(* IEC 61131-3 sources: 89152_FlorisHendrix_AfstudeerProject/89152_FlorisHendrix_ExamenProject/Stations/MachineControl/MachineControl/Class/VaranManager (part 5) *)

                DPRAM_Used.Total  += TempMem;
                DOCounter.Total   += 1;

            VARAN_CMD_CONTROL_WRITE,
            VARAN_CMD_MEMORY_WRITE:     // Write DO -------------------------------------------------------------------------------------------------------------------------------
                //32 Byte (Header) + 6 Byte (1 Byte Cmd, 4 Byte Addr, 1 Byte Len) + 1 Byte (Response) + n Byte (load data write) + 0 to 3 Byte (compensate missalignment)
                  TempMem := 32 + 6 + 1 + ud_WriteLength;
                  if (TempMem MOD 4) then
                    TempMem := TempMem + (4 - (TempMem MOD 4)); //increase memory, up to a value, which could be divided by 4
                  end_if;

                  case ud_DolType AND (NOT (VARAN_DOL_NOT_INSERT_DO_INTO_DOL)) of
                  // **************************************************
                    VARAN_DOL_DA:
                                  DPRAM_Used.DA_Wr    += TempMem;
                                  DOCounter.DA_Wr     += 1;
                  // **************************************************
                    VARAN_DOL_ISO:
                                  DPRAM_Used.ISO_Wr   += TempMem;
                                  DOCounter.ISO_Wr    += 1;
                  // **************************************************
                    VARAN_DOL_ASY:
                                  DPRAM_Used.ASY_Wr   += TempMem;
                                  DOCounter.ASY_Wr    += 1;
                  // **************************************************
                    VARAN_DOL_ADMIN:
                                  DPRAM_Used.Admin_Wr += TempMem;
                                  DOCounter.Admin_Wr  += 1;
                  // **************************************************
                    VARAN_DOL_IRQ:
                                  DPRAM_Used.IRQ_Wr   += TempMem;
                                  DOCounter.IRQ_Wr    += 1;
                  end_case;

                  DPRAM_Used.Total  += TempMem;
                  DOCounter.Total   += 1;

            VARAN_CMD_CONTROL_READ_WRITE,
            VARAN_CMD_MEMORY_READ_WRITE:// Read/Write DO -------------------------------------------------------------------------------------------------------------------------------
                  //32 Byte (Header) + 11 Byte (1 Byte Cmd, 4 Byte RdAddr, 1 Byte RdLen, 4 Byte WrAddr, 1 Byte WrLen) + 1 Byte (Response) + n Byte (load data read) + n Byte (load data write) + 0 to 3 Byte (compensate missalignment)
                  TempMem := 32 + 11 + 1 + ud_ReadLength + ud_WriteLength;
                  if (TempMem MOD 4) then
                    TempMem := TempMem + (4 - (TempMem MOD 4)); //increase memory, up to a value, which could be divided by 4
                  end_if;

                  case ud_DolType AND (NOT (VARAN_DOL_NOT_INSERT_DO_INTO_DOL)) of
                  // **************************************************
                    VARAN_DOL_DA:
                                  DPRAM_Used.DA_RdWr    += TempMem;
                                  DOCounter.DA_RdWr     += 1;
                  // **************************************************
                    VARAN_DOL_ISO:
                                  DPRAM_Used.ISO_RdWr   += TempMem;
                                  DOCounter.ISO_RdWr    += 1;
                  // **************************************************
                    VARAN_DOL_ASY:
                                  DPRAM_Used.ASY_RdWr   += TempMem;
                                  DOCounter.ASY_RdWr    += 1;
                  // **************************************************
                    VARAN_DOL_ADMIN:
                                  DPRAM_Used.Admin_RdWr += TempMem;
                                  DOCounter.Admin_RdWr  += 1;
                  // **************************************************
                    VARAN_DOL_IRQ:
                                  DPRAM_Used.IRQ_RdWr   += TempMem;
                                  DOCounter.IRQ_RdWr    += 1;
                  end_case;

                  DPRAM_Used.Total  += TempMem;
                  DOCounter.Total   += 1;

        end_case;

      end_if; // +++++++++++++++++++++++++++++++++++++++++++++++++++++++++++++++++++++++++++++++++++++++++++++++++++++++++++++++++++++++++++++++++++++++++++++++++++++++++++++++++++++++++++++++++

    end_if;
  else
    sd_retval := -100;	//Manager is off
  end_if;
END_FUNCTION

FUNCTION VaranManager::AddPayloadMoveDO
  VAR_INPUT
    p_ud_DoHandle 	                : ^UDINT;
    ud_bDoRequired 	                : UDINT;
    ud_DolType 	                    : UDINT;
    ud_Priority 	                  : UDINT;
    ud_PrescalerCounterThreshold 	  : UDINT;
    ud_PrescalerCounterStartValue 	: UDINT;
    ud_hSourceReadDoHandle 	        : UDINT;
    ud_ReadOffset 	                : UDINT;
    ud_hDestinationWriteDoHandle 	  : UDINT;
    ud_WriteOffset 	                : UDINT;
    ud_MoveDataLength 	            : UDINT;
  END_VAR
  VAR_OUTPUT
    sd_retval 	                    : DINT;
  END_VAR

#ifdef VM_DEBUG_PAYLOAD
  if b_PayloadSupport = false then
    // This method is not suppored without payload
    ((0)$^USINT)^ := 0;
  end_if;
#endif

  //look if we must execute Cyclic DOL list
  if ( ud_DolType = VARAN_DOL_ASY ) then
    s_CyHandles.b_ExecuteDOL := TRUE;			//set flag to execut Dol list
  end_if;

  sd_retval := MULTI_VARAN_iAddMoveDo(  phDoHandle                    := p_ud_DoHandle
                                      , bDoRequired                   := ud_bDoRequired
                                      , udDolType                     := ud_DolType
                                      , udPriority                    := ud_Priority
                                      , udPrescalerCounterThreshold   := ud_PrescalerCounterThreshold
                                      , udPrescalerCounterStartValue  := ud_PrescalerCounterStartValue
                                      , hSourceReadDoHandle           := ud_hSourceReadDoHandle
                                      , udReadOffset                  := ud_ReadOffset
                                      , hDestinationWriteDoHandle     := ud_hDestinationWriteDoHandle
                                      , udWriteOffset                 := ud_WriteOffset
                                      , udMoveDataLength              := ud_MoveDataLength
                                      );
  //look if an error occured
  if ( sd_retval <> VARANMANAGER_OK ) then
    s_ErrorVaranManager.f_AddRdDO := SetVaranDOError( sd_Error      := sd_retval
                                                    , b_manager_off := TRUE
                                                    , b_log         := TRUE
                                                    );
  else
    // Payload Move DO Mem Calculation
    if ( ud_DolType = VARAN_DOL_ASY ) then
      DPRAM_Used.ASY_Mov          += sizeof(LSL_VARANFRAMEPAYLOADMOVEHEADER);
      DPRAM_Used_Payload.ASY_Rd   += 1; // 1 Byte status
      DPRAM_Used_Payload.ASY_Wr   += sizeof(LSL_VARANFRAMEMOVEWRITEPAYLOAD);
      DOCounter.ASY_Mov           += 1;
    else
      DPRAM_Used.ISO_Mov          += sizeof(LSL_VARANFRAMEPAYLOADMOVEHEADER);
      DPRAM_Used_Payload.ISO_Rd   += 1; // 1 Byte status
      DPRAM_Used_Payload.ISO_Wr   += sizeof(LSL_VARANFRAMEMOVEWRITEPAYLOAD);
      DOCounter.ISO_Mov           += 1;
    end_if;

    DPRAM_Used.Total              += sizeof(LSL_VARANFRAMEPAYLOADMOVEHEADER) + 1 + sizeof(LSL_VARANFRAMEMOVEWRITEPAYLOAD);  // Header + Read Statusbyte + Write Payload
    DPRAM_Used_Payload.Total      += 1 + sizeof(LSL_VARANFRAMEMOVEWRITEPAYLOAD);  // Read Statusbyte + Write Payload
    DOCounter.Total               += 1;
  end_if;

END_FUNCTION

FUNCTION VaranManager::GetDataPointers
  VAR_INPUT
    ud_hDoHandle 	: UDINT;
    pp_ReadData 	: ^pVoid;
    pp_WriteData 	: ^pVoid;
  END_VAR
  VAR_OUTPUT
    sd_retval 	  : DINT;
  END_VAR

#ifdef VM_DEBUG_PAYLOAD
  if b_PayloadSupport = false then
    // This method is not suppored without payload
    ((0)$^USINT)^ := 0;
  end_if;
#endif

  // if there is no VARAN Interface available, we would crash at the call
  if pMultiVaran = NIL then
    sd_retval := VARANMANAGER_DRIVER_NOT_EXISTS;
    return;
  end_if;

  sd_retval :=  MULTI_VARAN_iGetDataPointers( hDoHandle   := ud_hDoHandle
                                            , ppvReadData := pp_ReadData
                                            , ppvWriteData:= pp_WriteData
                                            );

END_FUNCTION

FUNCTION VaranManager::GetModuleHandle
  VAR_INPUT
    p_us_PositionInfo 	: ^USINT;
    p_ud_ModuleHandle 	: ^UDINT;
  END_VAR
  VAR_OUTPUT
    sd_retval 	        : DINT;
  END_VAR

  // if there is no VARAN Interface available, we would crash at the call
  if pMultiVaran = NIL then
    sd_retval := VARANMANAGER_DRIVER_NOT_EXISTS;
    return;
  end_if;

  sd_retval := MULTI_VARAN_iGetNodeHandle(  udManagerNumber := VaranManagerNr
                                          , pszHardwarePath := p_us_PositionInfo
                                          , phNodeHandle    := p_ud_ModuleHandle
                                          );

END_FUNCTION

FUNCTION VaranManager::AddObjectCallback
	VAR_INPUT
		p_us_position_info 	: ^USINT;
		ud_action_ptr 	    : UDINT;
		ud_thisp 	          : UDINT;
		sd_required 	      : DINT;
	END_VAR
	VAR_OUTPUT
		sd_retval 	        : DINT;
	END_VAR
  VAR
    ud_NodeHandle       : UDINT;
  END_VAR

  if State = _NoVaranInterface then
    sd_retval := -100;
    return;
  end_if;
  //get right required flag
  if ( sd_required ) then
    sd_required := VARAN_DEVICE_REQUIRED;
  else
    sd_required := VARAN_DEVICE_DEFAULT;
  end_if;

  if b_PayloadSupport &
       pMultiVaran^.udVersion >= VM_MULTIVARAN_VERSION_FULL_PAYLOAD_AVAILABLE  then
    sd_retval := MULTI_VARAN_iGetNodeHandle ( udManagerNumber := VaranManagerNr
                                            , pszHardwarePath := p_us_position_info
                                            , phNodeHandle    := #ud_NodeHandle
                                            );

    if sd_retval <> VARANMANAGER_OK then
      return;
    end_if;

    //call OS - function to set callback
    sd_retval := MULTI_VARAN_iSetApplicationCallback( hNodeHandle           := ud_NodeHandle
                                                    , pfApplicationCallback := ud_action_ptr$pvoid
                                                    , pvUserData            := ud_thisp$pvoid
                                                    , udRequired            := sd_required$UDINT
                                                    );

  elsif pVaran then

    //call OS - function to set callback
    sd_retval := VARAN_iSetObjectCallback	( uiManager   := VaranManagerNr
                                          , pucNode     := p_us_position_info
                                          , uiCallback  := ud_action_ptr
                                          , uiThis      := ud_thisp
                                          , uiRequired  := sd_required$UDINT
                                          );
  end_if;

  //look for an error
  if ( sd_retval <> VARANMANAGER_OK ) then
    s_ErrorVaranManager.f_SetObjectCallback := SetVaranDOError	( sd_Error 		  := sd_retval
                                                                , b_manager_off	:= TRUE
                                                                , b_log			    := TRUE
                                                                );
  end_if;

END_FUNCTION

FUNCTION VaranManager::GetSPIDataFromID
	VAR_INPUT
		p_us_position_info 	: ^USINT;
		udListID 	          : UDINT;
		pData 	            : ^CHAR;
		udRequDataLength 	  : UDINT;
		pIDHeader 	        : ^t_s_SPIListHeader;
		udOffset 	          : UDINT;(* := 16#00 *)
	END_VAR
	VAR_OUTPUT
		sd_retval 	        : DINT;
	END_VAR
  VAR
    BaseListAddress     : UDINT;
    a_data              : ARRAY[0..31] OF UDINT;
  END_VAR

  if p_us_position_info & pData & udRequDataLength > 0 then

    //check OS version
    if ( _RTOSVersion < VM_SPI_OS_VERSION ) then
      // access of SPI flash not possible
      sd_retval := -2;
      return;
    end_if;

    // check if list is available and get size and offset in SPI flash
    if ( SearchSPIList(p_us_position_info, udListID, #BaseListAddress) <> VARANMANAGER_OK ) then
      sd_retval := -3;
      return;
    end_if;

    //read header of list
    sd_retval := ReadSPIDataComfort(p_us_position_info  := p_us_position_info,
                                    ud_offset           := BaseListAddress,
                                    ud_length	          := sizeof(t_s_SPIListHeader),
                                    p_data	            := ( #a_data )$^USINT
                                    );

    _memcpy(ptr1:=pIDHeader, ptr2:=#a_data[0], cntr:=sizeof(t_s_SPIListHeader));

    //look for an error and check if length is > 0
    if ( sd_retval <> VARANMANAGER_OK ) | ( a_data[ 2 ] = 0 ) then
      sd_retval := -4;
      return;
    end_if;

    //read the whole serial number string
    sd_retval := ReadSPIDataComfort( p_us_position_info := p_us_position_info,
                                     ud_offset	        := BaseListAddress + sizeof(t_s_SPIListHeader) + udOffset,  //+12 ist List Header
                                     ud_length	        := udRequDataLength,
                                     p_data		          := pData
                                    );

    //look for an error
    if ( sd_retval <> VARANMANAGER_OK ) then
      sd_retval := -5;
      return;
    end_if;
  else
    // invalid parameters
    sd_retval := -1;
  end_if;

END_FUNCTION

FUNCTION GLOBAL VaranManager::RaiseManagerError
	VAR_INPUT
		udReason 	: UDINT;
	END_VAR

  State := udReason$t_e_VaranErrors;

  if b_PayloadSupport & pMultiVaran^.udVersion >= VM_MULTIVARAN_VERSION_FULL_PAYLOAD_AVAILABLE  then
    MULTI_VARAN_iReportVaranError( diErrorNumber := udReason$DINT
                                 , hErrorNode    := vmNodeHandle
                                 );

  elsif pVaran & (pVaran^.udVersion >= 16#00001104 ) then
    VARAN_iSetManagerError( VaranManagerNr, udReason );
  end_if;

END_FUNCTION

FUNCTION VaranManager::GetExtNodeInfoDirectly
	VAR_INPUT
		pPara 	: ^t_VM_CMD_GetExtNodeInfo;
	END_VAR
	VAR_OUTPUT
		sd_retval 	: DINT;
	END_VAR
  VAR
    BaseListAddress     : UDINT;
    FoundIt             : BOOL;
    DataObjList         : ARRAY[0..31] OF UDINT;
    i                   : UDINT;
    sSPIListHeader      : t_s_SPIListHeader;
    sSPIIDList          : t_s_SPIIDListContent;
  END_VAR

  // initialize the retcode with error
  sd_retval := -1000;

  // the position info and pointer to the serial number are obligatory (always get the serial number)
  if pPara^.p_PositionInfo & pPara^.p_SerNoStr then

    //check OS version
    if ( _RTOSVersion < VM_SPI_OS_VERSION ) then
      // access of SPI flash not possible
      sd_retval := -1011;
      return;
    end_if;

    //************** GET THE ID LIST **********************************************

    //read SPI data
    sd_retval := ReadSPIData( p_us_position_info	:= pPara^.p_PositionInfo
                            , ud_offset				    := 0
                            , ud_length				    := 128 or VM_SPI_IDENT_LIST
                            , p_data				      := ( #DataObjList )$^USINT
                            );

    //look for an error
    if ( sd_retval <> VARANMANAGER_OK ) then
      sd_retval := -1010;
      return;
    end_if;

    //look for right Identifier
    if ( DataObjList[ 0 ] <> 16#12345678 ) then
      sd_retval := -1009;
      return;
    end_if;

    //look for valid length	(we only read 128 Byte at the moment [16Byte are header])
    if( DataObjList[ 3 ] > (128 - 16 ) ) then
      sd_retval := -1008;
      return;
    end_if;

    //************** GET THE SERIAL NUMBER ****************************************

    FoundIt := FALSE;

    //search for SPI Flash Configuration
    for i := 0 to DataObjList[ 3 ] / sizeof( UDINT ) do

      //look for configuration id in 3rd byte
      if ( ( DataObjList[ i + 4 ] and 16#FF00_0000 ) = VM_SPI_SERIALNO_ID ) then
        BaseListAddress := DataObjList[ i + 4 ] and 16#00FF_FFFF;
        FoundIt := TRUE;
      end_if;

    end_for;

    //if no entry is found
    if FoundIt = FALSE then
      sd_retval := -1007;
      return;
    end_if;

    //read header of serial number list
    sd_retval := ReadSPIDataComfort(p_us_position_info  := pPara^.p_PositionInfo,
                                    ud_offset           := BaseListAddress,
                                    ud_length	          := sizeof(t_s_SPIListHeader),
                                    p_data	            := ( #sSPIListHeader )$^USINT
                                   );

    //look for an error and check if length is > 0 and smaller than max length
    if ( sd_retval <> VARANMANAGER_OK ) | ( sSPIListHeader.ListLength = 0 ) | ( sSPIListHeader.ListLength > SERNO_STRING_SIZE ) then
      sd_retval := -1006;
      return;
    end_if;

    //read the whole serial number string
    sd_retval := ReadSPIDataComfort( p_us_position_info := pPara^.p_PositionInfo,
                                     ud_offset	        := BaseListAddress + sizeof(t_s_SPIListHeader),
                                     ud_length	        := sSPIListHeader.ListLength,
                                     p_data		          := pPara^.p_SerNoStr
                                   );

    //add string termination
    (pPara^.p_SerNoStr + sSPIListHeader.ListLength)^ := 0;

    //look for an error
    if ( sd_retval <> VARANMANAGER_OK ) then
      sd_retval := -1005;
      return;
    end_if;

      //************** GET THE HARDWARE VERSION AND LICENSE NUMBER ******************

    // check if any additional data is needed
    if pPara^.p_HwVersion | pPara^.p_LicenseNo then

      FoundIt := FALSE;

      //search for SPI Flash Configuration
      for i := 0 to DataObjList[ 3 ] / sizeof( UDINT ) do

        //look for configuration id in 3rd byte
        if ( ( DataObjList[ i + 4 ] and 16#FF00_0000 ) = VM_SPI_IDENTIFICATION_LIST ) then
          BaseListAddress := DataObjList[ i + 4 ] and 16#00FF_FFFF;
          FoundIt := TRUE;
        end_if;

      end_for;

      //if no entry found
      if FoundIt = FALSE then
        sd_retval := -1004;
        return;
      end_if;

      //read header of identification list
      sd_retval := ReadSPIDataComfort(p_us_position_info  := pPara^.p_PositionInfo,
                                      ud_offset           := BaseListAddress,
                                      ud_length	          := sizeof(t_s_SPIListHeader),
                                      p_data	            := ( #sSPIListHeader )$^USINT
                                     );

      //look for an error and check if length is >= 16 (hw version is at offset 12 with 4 bytes)
      if ( sd_retval <> VARANMANAGER_OK ) | ( sSPIListHeader.ListLength < 16 ) then
        sd_retval := -1003;
        return;
      end_if;

      //read the hardware version
      sd_retval := ReadSPIDataComfort( p_us_position_info := pPara^.p_PositionInfo,
                                       ud_offset	        := BaseListAddress + sizeof(t_s_SPIListHeader),
                                       ud_length	        := sizeof(t_s_SPIIDListContent),
                                       p_data		          := (#sSPIIDList)$^USINT
                                     );

      //look for an error
      if ( sd_retval <> VARANMANAGER_OK ) then
        sd_retval := -1002;
        return;
      end_if;

      // if the HwVersion pointer is valid => store the HwVersion there
      if pPara^.p_HwVersion then
        pPara^.p_HwVersion^ := sSPIIDList.HwVersion;
      end_if;

      // if the LicenseNo pointer is valid => store the HwVersion there
      if pPara^.p_LicenseNo then
        pPara^.p_LicenseNo^ := sSPIIDList.LicenseNo;
      end_if;
    end_if;

    // success
    sd_retval := 0;
  else
    // invalid parameters
    sd_retval := -1001;
  end_if;

END_FUNCTION
